(* IEC 61131-3 sources: kns-port-domestic/upstream/kns-pump-station/src/POUs/Log/FB_EventLog, 15 files *)

(* ---- FB_EventLog.decl.st ---- *)
// Назначение: журнал событий КНС-1 — кольцевой буфер LOG_CAPACITY (200) записей ST_EventRecord в ОЗУ:
//             переходы тревог устройств, станции и LIC101 (приёмник PL.I_AlarmSink, ссылка в
//             PL.GVL_Lib.itfAlarmSink) и события станции (I_StationEventSink, номер STN_EVENT_ID_BASE + код).
//             При переполнении затирается самая старая запись (udiOverwritten). Метки: UTC от
//             SysTimeRtcHighResGet (мс; 0 — часы недоступны) и время процесса lrMono_s по itfTime.
//             Страница HMI (FillView), курсор внешних клиентов (FillFeed), снимок для CSV (TakeSnapshot —
//             MainTask, GetSnapshotRecord — SlowTask). Тело пустое: записи делают методы в момент события.
// Автор:      kr0nsch
// Версия:     0.1.0
// Документ:   docs/DESIGN.md, раздел 9.1; docs/04_algorithms.md, раздел 16
FUNCTION_BLOCK FB_EventLog IMPLEMENTS PL.I_AlarmSink, I_StationEventSink
VAR_INPUT
    itfTime : PL.I_TimeSource;      // GVL_Time.fbClockMain (присваивает PRG_Station каждый цикл); 0 — LTIME()
END_VAR
VAR_OUTPUT
    uiCount        : UINT;          // записей в кольце, 0…LOG_CAPACITY
    udiSeqLast     : UDINT;         // номер последней записи; 0 — записей не было
    udiOverwritten : UDINT;         // затёрто записей с запуска
    xClockValid    : BOOL;          // последняя запись: RTC ответил и время правдоподобно
END_VAR
VAR
    astRing     : ARRAY[0..GVL_Const.LOG_CAPACITY - 1] OF ST_EventRecord;   // кольцо
    uiHead      : UINT;             // индекс следующей записи в кольце
    astSnapshot : ARRAY[0..GVL_Const.LOG_CAPACITY - 1] OF ST_EventRecord;   // снимок, от старой записи к новой
    uiSnapCount : UINT;             // записей в снимке
    fbSysTime   : PL.FB_SystemTime; // источник времени без itfTime
END_VAR

(* ---- FillFeed.method.decl.st ---- *)
// Курсор внешнего клиента: до LOG_FEED_ROWS записей от номера MAX(stFeed.udiFromSeq, самая старая) к новым.
// udiFromSeq < udiSeqFirst — клиент пропустил затёртые записи (видит по номерам)
METHOD FillFeed
VAR_IN_OUT
    stFeed : ST_EventFeed;          // GVL_Log.stEventFeed
END_VAR
VAR
    udiSeq  : UDINT;                // номер записи очередной строки
    uiRow   : UINT;                 // строка курсора
    stEmpty : ST_EventRecord;       // пустая строка
END_VAR

(* ---- FillFeed.method.impl.st ---- *)
stFeed.udiSeqLast := udiSeqLast;
stFeed.udiSeqFirst := udiSeqLast + 1 - UINT_TO_UDINT(uiCount);
stFeed.wReserve := 0;
udiSeq := MAX(stFeed.udiFromSeq, stFeed.udiSeqFirst);
stFeed.uiCount := 0;
FOR uiRow := 1 TO GVL_Const.LOG_FEED_ROWS DO
    IF udiSeq <= udiSeqLast THEN
        // udiSeqLast - udiSeq < uiCount <= LOG_CAPACITY: возраст помещается в UINT
        GetRecord(uiAge := UDINT_TO_UINT(udiSeqLast - udiSeq), stRecord => stFeed.astRow[uiRow]);
        stFeed.uiCount := uiRow;
        udiSeq := udiSeq + 1;
    ELSE
        stFeed.astRow[uiRow] := stEmpty;
    END_IF
END_FOR

(* ---- FillView.method.decl.st ---- *)
// Страница журнала для HMI: номер страницы stView.uiPage (0 — новые) ограничивается последней страницей,
// строки — новые сверху; строки после последней записи — пустые (udiSeq = 0)
METHOD FillView
VAR_IN_OUT
    stView : ST_EventView;          // GVL_Log.stEventView
END_VAR
VAR
    uiRow      : UINT;              // строка страницы
    uiAgeFirst : UINT;              // возраст записи первой строки
END_VAR

(* ---- FillView.method.impl.st ---- *)
stView.uiCount := uiCount;
stView.uiPageCount := MAX(1, (uiCount + GVL_Const.LOG_VIEW_ROWS - 1) / GVL_Const.LOG_VIEW_ROWS);
IF stView.uiPage >= stView.uiPageCount THEN
    stView.uiPage := stView.uiPageCount - 1;
END_IF
stView.wReserve := 0;
uiAgeFirst := stView.uiPage * GVL_Const.LOG_VIEW_ROWS;
FOR uiRow := 1 TO GVL_Const.LOG_VIEW_ROWS DO
    GetRecord(uiAge := uiAgeFirst + uiRow - 1, stRecord => stView.astRow[uiRow]);
END_FOR

(* ---- GetRecord.method.decl.st ---- *)
// Запись по возрасту: 0 — самая новая; FALSE — такой записи нет (stRecord — нули, udiSeq = 0)
METHOD GetRecord : BOOL
VAR_INPUT
    uiAge : UINT;                   // 0 — новая, uiCount - 1 — самая старая
END_VAR
VAR_OUTPUT
    stRecord : ST_EventRecord;
END_VAR
VAR
    stEmpty : ST_EventRecord;       // пустая запись
END_VAR

(* ---- GetRecord.method.impl.st ---- *)
IF uiAge < uiCount THEN
    // uiAge < uiCount <= LOG_CAPACITY: индекс не уходит в минус
    stRecord := astRing[(uiHead + GVL_Const.LOG_CAPACITY - 1 - uiAge) MOD GVL_Const.LOG_CAPACITY];
    GetRecord := TRUE;
ELSE
    stRecord := stEmpty;
    GetRecord := FALSE;
END_IF

(* ---- GetSnapshotRecord.method.decl.st ---- *)
// Запись снимка (SlowTask): 0 — самая старая; FALSE — индекс вне снимка (stRecord — нули)
METHOD GetSnapshotRecord : BOOL
VAR_INPUT
    uiIndex : UINT;                 // 0…SnapshotCount - 1
END_VAR
VAR_OUTPUT
    stRecord : ST_EventRecord;
END_VAR
VAR
    stEmpty : ST_EventRecord;       // пустая запись
END_VAR

(* ---- GetSnapshotRecord.method.impl.st ---- *)
IF uiIndex < uiSnapCount THEN
    stRecord := astSnapshot[uiIndex];
    GetSnapshotRecord := TRUE;
ELSE
    stRecord := stEmpty;
    GetSnapshotRecord := FALSE;
END_IF

(* ---- LogEvent.method.decl.st ---- *)
// I_StationEventSink: событие станции — запись вида Station с номером STN_EVENT_ID_BASE + код, приоритетом
// None и состояниями Normal; TRUE — записано
METHOD LogEvent : BOOL
VAR_INPUT
    eEvent : E_StationEvent;        // номер записи = STN_EVENT_ID_BASE + eEvent
    rValue : REAL;                  // аргумент (номер насоса, параметра, строк…)
END_VAR

(* ---- OnAlarmEvent.method.decl.st ---- *)
// PL.I_AlarmSink: переход тревоги (PL.FB_Alarm устройств, станции, LIC101) — запись вида Alarm; всегда TRUE
METHOD OnAlarmEvent : BOOL
VAR_IN_OUT CONSTANT
    stEvent : PL.ST_AlarmEvent;     // событие
END_VAR

(* ---- Store.method.decl.st ---- *)
// Добавить запись: сквозной номер, метки UTC и времени процесса; в полном кольце затирается самая старая.
// Всегда TRUE: кольцо не переполняется
METHOD PRIVATE Store : BOOL
VAR_INPUT
    eKind     : E_EventKind;
    ePriority : PL.E_AlarmPriority;
    udiId     : UDINT;
    eOldState : PL.E_AlarmState;
    eNewState : PL.E_AlarmState;
    eReason   : PL.E_AlarmEventReason;
    rValue    : REAL;
END_VAR
VAR
    uliUtc_ms  : ULINT;             // ответ часов реального времени
    itfTimeAct : PL.I_TimeSource;   // действующий источник времени процесса
END_VAR

(* ---- Store.method.impl.st ---- *)
itfTimeAct := itfTime;
IF itfTimeAct = 0 THEN
    itfTimeAct := fbSysTime;
END_IF
// часы реального времени: ошибка или время раньше LOG_UTC_MIN_MS (часы не выставлены) — метка 0
uliUtc_ms := F_UtcNowMs();
xClockValid := uliUtc_ms <> 0;
udiSeqLast := udiSeqLast + 1;
astRing[uiHead].udiSeq := udiSeqLast;
astRing[uiHead].eKind := eKind;
astRing[uiHead].ePriority := ePriority;
astRing[uiHead].udiId := udiId;
astRing[uiHead].eOldState := eOldState;
astRing[uiHead].eNewState := eNewState;
astRing[uiHead].eReason := eReason;
astRing[uiHead].wReserve := 0;
astRing[uiHead].rValue := rValue;
astRing[uiHead].uliUtc_ms := uliUtc_ms;
astRing[uiHead].lrMono_s := PL.F_LTimeToSec(ltIn := itfTimeAct.Now());
uiHead := (uiHead + 1) MOD GVL_Const.LOG_CAPACITY;
IF uiCount < GVL_Const.LOG_CAPACITY THEN
    uiCount := uiCount + 1;
ELSE
    udiOverwritten := udiOverwritten + 1;
END_IF
Store := TRUE;

(* ---- TakeSnapshot.method.decl.st ---- *)
// Снимок кольца для выгрузки CSV (MainTask): записи от старой к новой в astSnapshot. TRUE — снимок сделан.
// Вызывать, только пока SlowTask не пишет файл (GVL_Log.eExportState не Writing): снимок читает SlowTask
METHOD TakeSnapshot : BOOL
VAR
    uiI : UINT;                     // номер записи снимка, с 1
END_VAR

(* ---- TakeSnapshot.method.impl.st ---- *)
uiSnapCount := uiCount;
FOR uiI := 1 TO uiSnapCount DO
    GetRecord(uiAge := uiSnapCount - uiI, stRecord => astSnapshot[uiI - 1]);
END_FOR
TakeSnapshot := TRUE;
